//{attribute 'Tc2GvlVarNames'}
VAR_GLOBAL PERSISTENT
	Errors: DINT;
	SetSlaveToOP_ON     : BOOL:=TRUE;
	bEnableAutoResetEncoder: BOOL:=TRUE;
END_VAR

(* stored: Version 1.1.0.1, ProductVersion 3.1.4024.13
   GVL Global_Persistent: Id {3d408214-16c8-4d4c-9564-6c4ba0d62286} *)
